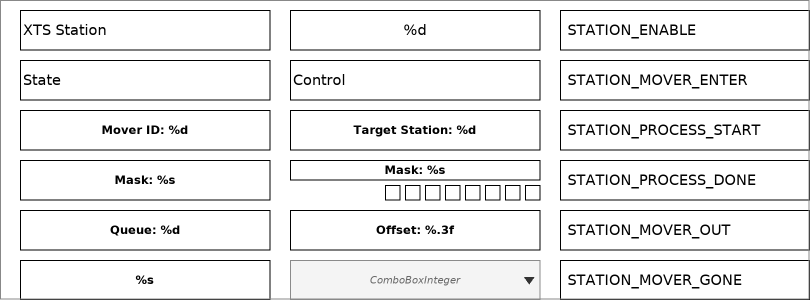
VISUALIZATION STATION_VISU  // 810x300
    Rectangle (20,10 250x40), "XTS Station"
    Rectangle (290,10 250x40), "%d", text variable: VISU_POOL.nStationSelected
        OnMouseClick: write the text variable via VisuDialogs.Numpad, min 1, max MAX_STATION, title 'Selected Station'
    Rectangle (20,60 250x40), "State"
    Rectangle (290,60 250x40), "Control"
    Rectangle (20,210 250x40), "Queue: %d", text variable: GVL_XTS.StationState[VISU_POOL.nStationSelected].nQueue
    Rectangle (20,110 250x40), "Mover ID: %d", text variable: GVL_XTS.StationState[VISU_POOL.nStationSelected].nMoverId
    Rectangle (20,160 250x40), "Mask: %s", text variable: GVL_APPLICATION.VisuPoolData.sStationStateMask
    Rectangle (20,260 250x40), "%s", text variable: GVL_APPLICATION.VisuPoolData.sStationState
    ComboBoxInteger (290,260 250x40), variable: GVL_XTS.StationCtrl[VISU_POOL.nStationSelected].eCmd, text list: 'TL_E_CTRL_STATION'
    Rectangle (290,210 250x40), "Offset: %.3f", text variable: GVL_XTS.StationCtrl[VISU_POOL.nStationSelected].rOffset
    Rectangle (290,110 250x40), "Target Station: %d", text variable: GVL_XTS.StationCtrl[VISU_POOL.nStationSelected].nTargetStation
        OnMouseClick: write the text variable via VisuDialogs.Numpad, min 1, max MAX_STATION, title 'Target Station'
    Rectangle (290,160 250x20), "Mask: %s", text variable: GVL_APPLICATION.VisuPoolData.sStationCtrlMask
    Rectangle (525,185 15x15)
        toggle GVL_XTS.StationCtrl[VISU_POOL.nStationSelected].nMask.0
    Rectangle (505,185 15x15)
        toggle GVL_XTS.StationCtrl[VISU_POOL.nStationSelected].nMask.1
    Rectangle (485,185 15x15)
        toggle GVL_XTS.StationCtrl[VISU_POOL.nStationSelected].nMask.2
    Rectangle (465,185 15x15)
        toggle GVL_XTS.StationCtrl[VISU_POOL.nStationSelected].nMask.3
    Rectangle (445,185 15x15)
        toggle GVL_XTS.StationCtrl[VISU_POOL.nStationSelected].nMask.4
    Rectangle (425,185 15x15)
        toggle GVL_XTS.StationCtrl[VISU_POOL.nStationSelected].nMask.5
    Rectangle (405,185 15x15)
        toggle GVL_XTS.StationCtrl[VISU_POOL.nStationSelected].nMask.6
    Rectangle (385,185 15x15)
        toggle GVL_XTS.StationCtrl[VISU_POOL.nStationSelected].nMask.7
    Rectangle (560,10 250x40), "STATION_ENABLE", colour toggle: GVL_APPLICATION.VisuPoolData.bStationEnable
        OnMouseClick: execute { GVL_XTS.StationCtrl[VISU_POOL.nMoverSelected].Cmd := E_STATION_CTRL.STATION_ENABLE; }
    Rectangle (560,60 250x40), "STATION_MOVER_ENTER", colour toggle: GVL_APPLICATION.VisuPoolData.bStationEnter
        OnMouseClick: execute { GVL_XTS.StationCtrl[VISU_POOL.nMoverSelected].Cmd := E_STATION_CTRL.STATION_MOVER_ENTER; }
    Rectangle (560,110 250x40), "STATION_PROCESS_START", colour toggle: GVL_APPLICATION.VisuPoolData.bStationStart
        OnMouseClick: execute { GVL_XTS.StationCtrl[VISU_POOL.nMoverSelected].Cmd := E_STATION_CTRL.STATION_PROCESS_START; }
    Rectangle (560,160 250x40), "STATION_PROCESS_DONE", colour toggle: GVL_APPLICATION.VisuPoolData.bStationDone
        OnMouseClick: execute { GVL_XTS.StationCtrl[VISU_POOL.nMoverSelected].Cmd := E_STATION_CTRL.STATION_PROCESS_DONE; }
    Rectangle (560,210 250x40), "STATION_MOVER_OUT", colour toggle: GVL_APPLICATION.VisuPoolData.bStationOut
        OnMouseClick: execute { GVL_XTS.StationCtrl[VISU_POOL.nMoverSelected].Cmd := E_STATION_CTRL.STATION_MOVER_OUT; }
    Rectangle (560,260 250x40), "STATION_MOVER_GONE", colour toggle: GVL_APPLICATION.VisuPoolData.bStationGone
        OnMouseClick: execute { GVL_XTS.StationCtrl[VISU_POOL.nMoverSelected].Cmd := E_STATION_CTRL.STATION_MOVER_GONE; }
END_VISUALIZATION

(* stored: Version 1.1.0.1
   Visu STATION_VISU: Id {5611794e-4b72-4a4d-ad30-97e40a2b205b} *)
